(*
SPDX-FileCopyrightText: © 2026 Oleksandr Tiutyk <trofimich@gmail.com>
SPDX-License-Identifier: MIT
License: https://opensource.org/license/mit
*)

(*!
<summary>Mock root controller for automation component lifecycle and hierarchy tests.</summary>
*)

FUNCTION_BLOCK MockAutomationController EXTENDS TOF_Automation.AutomationController<0>
VAR_STAT
	{attribute 'hide'}
	_ClassName : STRING := __POUNAME();
END_VAR

PROPERTY Children : REFERENCE TO ARRAY [0.._ChildCount - 1] OF TOF_Automation.IChildAutomationComponent
GET
Children REF= 0;
END_GET
END_PROPERTY

{attribute 'monitoring' := 'call'}
PROPERTY ClassName : REFERENCE TO STRING
GET
ClassName REF= _ClassName;
END_GET
END_PROPERTY

METHOD FB_init : BOOL
VAR_INPUT
	bInitRetains : BOOL; // TRUE: the retain variables are initialized (reset warm / reset cold)
	bInCopyCode : BOOL;  // TRUE: the instance will be copied to the copy code afterward (online change)
	name : WSTRING;
END_VAR
END_METHOD

{attribute 'monitoring' := 'call'}
PROPERTY NamespaceName : REFERENCE TO STRING
GET
NamespaceName REF= CurrentNamespace.Name;
END_GET
END_PROPERTY

{attribute 'monitoring' := 'call'}
PROPERTY SelfSize : ULINT
GET
SelfSize := XSIZEOF(THIS^);
END_GET
END_PROPERTY

END_FUNCTION_BLOCK

(* stored: Version 1.1.0.1, ProductVersion 3.1.4026.21
   POU MockAutomationController: Id {b1387f91-0a12-44ed-8c2c-5c2ab7f18700}, SpecialFunc None
   Property Children: Id {fa890d89-8bdf-4ea5-8f9d-011c91dc1c3b}
   Get Get: Id {568c87d4-32ef-4f19-9ae0-c1f3d2b9f5d1}
   Property ClassName: Id {4013738d-e570-41bf-a39d-46cce17c11f7}
   Get Get: Id {9069a7f4-690e-413d-9ca5-71262b49a219}
   Method FB_init: Id {c78a8024-b95b-438b-a697-782c5f4b9636}
   Property NamespaceName: Id {b188574b-a97a-41b7-a9f2-a27c833cee31}
   Get Get: Id {70c14aa1-b4fb-4080-aeba-71551ae994a8}
   Property SelfSize: Id {e1f8d4e4-cadf-4f07-9eb1-4d1532dbb9c4}
   Get Get: Id {26e8ca1d-6bbc-4f27-a90d-bff3d9976c38} *)
